(* PLC project TBEN_L5_PLC11.project, CODESYS CODESYS V3.5 SP21 Patch 1 *)
(* stored: creationDateTime 2026-11-07T15:34:51.3235159, modificationDateTime 2026-11-07T15:09:07.4034196 *)

{attribute 'qualified_only'}
// Loại việc ISDU đang chạy trong FB_IolDevBase
TYPE E_IolDevJob :
(
    NONE     := 0,
    IDENT    := 1,  // đọc index 16..24
    PARAM_RD := 2,  // đọc 1 tham số trong bảng
    PARAM_WR := 3,  // ghi 1 tham số trong bảng
    CUSTOM   := 4   // ISDU tự do của lớp con (system command, event list...)
) INT;
END_TYPE
